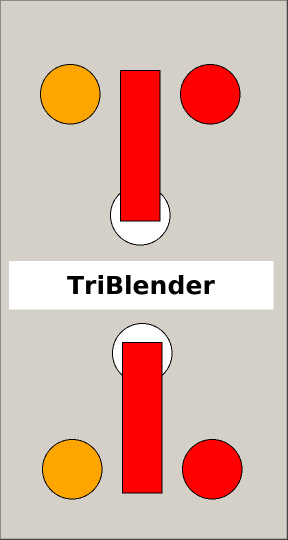
VISUALIZATION vis_TriBlenderPipe  // 288x540
    Rectangle (0,0 288x540)
    Ellipse (112,323 60x60)
        OnMouseClick: execute { eTriBlenderPipe_In:=E_TriBlenderPipe.eNone; }
    Ellipse (42,439 60x60)
        OnMouseClick: execute { eTriBlenderPipe_In:=E_TriBlenderPipe.eMarinada; }
    Ellipse (182,439 60x60)
        OnMouseClick: execute { eTriBlenderPipe_In:=E_TriBlenderPipe.eColor; }
    Ellipse (110,185 60x60)
        OnMouseClick: execute { eTriBlenderPipe_Out:=E_TriBlenderPipe.eNone; }
    Ellipse (40,64 60x60)
        OnMouseClick: execute { eTriBlenderPipe_Out:=E_TriBlenderPipe.eMarinada; }
    Ellipse (180,64 60x60)
        OnMouseClick: execute { eTriBlenderPipe_Out:=E_TriBlenderPipe.eColor; }
    RoundedRectangle (120,70 40x151), angle -30, invisible if: eTriBlenderPipe_Out<>E_TriBlenderPipe.eMarinada
        OnMouseClick: execute { eTriBlenderPipe_Out:=E_TriBlenderPipe.eNone; }
    RoundedRectangle (120,70 40x151), angle 30, invisible if: eTriBlenderPipe_Out<>E_TriBlenderPipe.eColor
        OnMouseClick: execute { eTriBlenderPipe_Out:=E_TriBlenderPipe.eNone; }
    RoundedRectangle (122,342 40x151), angle 30, invisible if: eTriBlenderPipe_In<>E_TriBlenderPipe.eMarinada
        OnMouseClick: execute { eTriBlenderPipe_In:=E_TriBlenderPipe.eNone; }
    RoundedRectangle (122,342 40x151), angle -30, invisible if: eTriBlenderPipe_In<>E_TriBlenderPipe.eColor
        OnMouseClick: execute { eTriBlenderPipe_In:=E_TriBlenderPipe.eNone; }
    Textfield (8,260 266x50), "TriBlender"
END_VISUALIZATION

(* stored: Version 1.1.0.1, ProductVersion 3.1.4024.12
   Visu vis_TriBlenderPipe: Id {c2ab4589-0e35-4b3d-a1ec-5e0f0c3193c6} *)
